// TIA Portal V20 export
VAR_GLOBAL   // PLC tag table "COGNEX_ETIKETA"
   "COG_ETIKETA_COG_ETIKETA_is3800-TriggerEnable" AT %Q2.0 : Bool;
   "COG_ETIKETA_COG_ETIKETA_is3800-Trigger" AT %Q2.1 : Bool;
   "COG_ETIKETA_is3800-ClearExposureComplete" AT %Q2.2 : Bool;
   "COG_ETIKETA_is3800-Set Offline" AT %Q2.7 : Bool;
   "COG_ETIKETA_is3800-TriggerReady" AT %I2.0 : Bool;
   "COG_ETIKETA_is3800-TriggerAck" AT %I2.1 : Bool;
   "COG_ETIKETA_is3800-ExposureComplete" AT %I2.2 : Bool;
   "COG_ETIKETA_is3800-AcquCOG_ETIKETA_isitionError" AT %I2.3 : Bool;
   "COG_ETIKETA_is3800-Offline Reason" AT %I2.4 : Bool;
   "COG_ETIKETA_is3800-Offline Reason(1)" AT %I2.5 : Bool;
   "COG_ETIKETA_is3800-Offline Reason(2)" AT %I2.6 : Bool;
   "COG_ETIKETA_is3800-Online" AT %I2.7 : Bool;
   "COG_ETIKETA_is3800-AcquCOG_ETIKETA_isitionID" AT %IW4 : Int;
   "COG_ETIKETA_is3800-BufferResultsEnable" AT %Q3.0 : Bool;
   "COG_ETIKETA_is3800-InspectionResultsAck" AT %Q3.1 : Bool;
   "COG_ETIKETA_is3800-SetUserData" AT %Q3.2 : Bool;
   "COG_ETIKETA_is3800-ExecuteCommand/JobLoad" AT %Q3.3 : Bool;
   "COG_ETIKETA_is3800-ClearError" AT %Q3.7 : Bool;
   "COG_ETIKETA_is3800-Reserved" AT %I10.0 : Bool;
   "COG_ETIKETA_is3800-InspectionCompleted" AT %I10.1 : Bool;
   "COG_ETIKETA_is3800-ResultsBufferOverrun" AT %I10.2 : Bool;
   "COG_ETIKETA_is3800-ResultsValid" AT %I10.3 : Bool;
   "COG_ETIKETA_is3800-CommandExecuting" AT %I10.4 : Bool;
   "COG_ETIKETA_is3800-CommandCompleted" AT %I10.5 : Bool;
   "COG_ETIKETA_is3800-CommandFailed" AT %I10.6 : Bool;
   "COG_ETIKETA_is3800-SetUserDataAck" AT %I10.7 : Bool;
   "COG_ETIKETA_is3800-ResultsPassed (Job)" AT %I11.0 : Bool;
   "COG_ETIKETA_is3800-SystemValidated" AT %I11.1 : Bool;
   "COG_ETIKETA_is3800-Error" AT %I11.7 : Bool;
   "COG_ETIKETA_is3800-ErrorCode" AT %IW12 : Word;
   "COG_ETIKETA_is3800-CommandID" AT %QW64 : Word;
   "COG_ETIKETA_is3800-Current Job ID" AT %IW68 : Word;
   "COG_ETIKETA_is3800-CommandResultCode" AT %IW70 : Word;
   "COG_ETIKETA_is3800-ExternalEvent[0]" AT %Q4.0 : Bool;
   "COG_ETIKETA_is3800-ExternalEvent[1]" AT %Q4.1 : Bool;
   "COG_ETIKETA_is3800-ExternalEvent[2]" AT %Q4.2 : Bool;
   "COG_ETIKETA_is3800-ExternalEvent[3]" AT %Q4.3 : Bool;
   "COG_ETIKETA_is3800-ExternalEvent[4]" AT %Q4.4 : Bool;
   "COG_ETIKETA_is3800-ExternalEvent[5]" AT %Q4.5 : Bool;
   "COG_ETIKETA_is3800-ExternalEvent[6]" AT %Q4.6 : Bool;
   "COG_ETIKETA_is3800-ExternalEvent[7]" AT %Q4.7 : Bool;
   "COG_ETIKETA_is3800-ExternalEventAck[0]" AT %I6.0 : Bool;
   "COG_ETIKETA_is3800-ExternalEventAck[1]" AT %I6.1 : Bool;
   "COG_ETIKETA_is3800-ExternalEventAck[2]" AT %I6.2 : Bool;
   "COG_ETIKETA_is3800-ExternalEventAck[3]" AT %I6.3 : Bool;
   "COG_ETIKETA_is3800-ExternalEventAck[4]" AT %I6.4 : Bool;
   "COG_ETIKETA_is3800-ExternalEventAck[5]" AT %I6.5 : Bool;
   "COG_ETIKETA_is3800-ExternalEventAck[6]" AT %I6.6 : Bool;
   "COG_ETIKETA_is3800-ExternalEventAck[7]" AT %I6.7 : Bool;
   "COG_ETIKETA_is3800-UserData[0]" AT %QB66 : Byte;
   "COG_ETIKETA_is3800-UserData[1]" AT %QB67 : Byte;
   "COG_ETIKETA_is3800-UserData[2]" AT %QB68 : Byte;
   "COG_ETIKETA_is3800-UserData[3]" AT %QB69 : Byte;
   "COG_ETIKETA_is3800-UserData[4]" AT %QB70 : Byte;
   "COG_ETIKETA_is3800-UserData[5]" AT %QB71 : Byte;
   "COG_ETIKETA_is3800-UserData[6]" AT %QB72 : Byte;
   "COG_ETIKETA_is3800-UserData[7]" AT %QB73 : Byte;
   "COG_ETIKETA_is3800-UserData[8]" AT %QB74 : Byte;
   "COG_ETIKETA_is3800-UserData[9]" AT %QB75 : Byte;
   "COG_ETIKETA_is3800-UserData[10]" AT %QB76 : Byte;
   "COG_ETIKETA_is3800-UserData[11]" AT %QB77 : Byte;
   "COG_ETIKETA_is3800-UserData[12]" AT %QB78 : Byte;
   "COG_ETIKETA_is3800-UserData[13]" AT %QB79 : Byte;
   "COG_ETIKETA_is3800-UserData[14]" AT %QB80 : Byte;
   "COG_ETIKETA_is3800-UserData[15]" AT %QB81 : Byte;
   "COG_ETIKETA_is3800-InspectionID" AT %IW72 : Word;
   "COG_ETIKETA_is3800-InspectionResultsCode" AT %IW74 : Int;
   "COG_ETIKETA_is3800-InspectionResults_0" AT %IB76 : Byte;
   "COG_ETIKETA_is3800-InspectionResults_1" AT %IB77 : Byte;
   "COG_ETIKETA_is3800-InspectionResults_2" AT %IB78 : Byte;
   "COG_ETIKETA_is3800-InspectionResults_3" AT %IB79 : Byte;
   "COG_ETIKETA_is3800-InspectionResults_4" AT %IB80 : Byte;
   "COG_ETIKETA_is3800-InspectionResults_5" AT %IB81 : Byte;
   "COG_ETIKETA_is3800-InspectionResults_6" AT %IB82 : Byte;
   "COG_ETIKETA_is3800-InspectionResults_7" AT %IB83 : Byte;
   "COG_ETIKETA_is3800-InspectionResults_8" AT %IB84 : Byte;
   "COG_ETIKETA_is3800-InspectionResults_9" AT %IB85 : Byte;
   "COG_ETIKETA_is3800-InspectionResults_10" AT %IB86 : Byte;
   "COG_ETIKETA_is3800-InspectionResults_11" AT %IB87 : Byte;
   "COG_ETIKETA_is3800-InspectionResults_12" AT %IB88 : Byte;
   "COG_ETIKETA_is3800-InspectionResults_13" AT %IB89 : Byte;
   "COG_ETIKETA_is3800-InspectionResults_14" AT %IB90 : Byte;
   "COG_ETIKETA_is3800-InspectionResults_15" AT %IB91 : Byte;
   "COG_ETIKETA_is3800-InspectionResults_16" AT %IB92 : Byte;
   "COG_ETIKETA_is3800-InspectionResults_17" AT %IB93 : Byte;
   "COG_ETIKETA_is3800-InspectionResults_18" AT %IB94 : Byte;
   "COG_ETIKETA_is3800-InspectionResults_19" AT %IB95 : Byte;
   "COG_ETIKETA_is3800-InspectionResults_20" AT %IB96 : Byte;
   "COG_ETIKETA_is3800-InspectionResults_21" AT %IB97 : Byte;
   "COG_ETIKETA_is3800-InspectionResults_22" AT %IB98 : Byte;
   "COG_ETIKETA_is3800-InspectionResults_23" AT %IB99 : Byte;
   "COG_ETIKETA_is3800-InspectionResults_24" AT %IB100 : Byte;
   "COG_ETIKETA_is3800-InspectionResults_25" AT %IB101 : Byte;
   "COG_ETIKETA_is3800-InspectionResults_26" AT %IB102 : Byte;
   "COG_ETIKETA_is3800-InspectionResults_27" AT %IB103 : Byte;
   "COG_ETIKETA_is3800-InspectionResults_28" AT %IB104 : Byte;
   "COG_ETIKETA_is3800-InspectionResults_29" AT %IB105 : Byte;
   "COG_ETIKETA_is3800-InspectionResults_30" AT %IB106 : Byte;
   "COG_ETIKETA_is3800-InspectionResults_31" AT %IB107 : Byte;
   "COG_ETIKETA_is3800-InspectionResults_32" AT %IB108 : Byte;
   "COG_ETIKETA_is3800-InspectionResults_33" AT %IB109 : Byte;
   "COG_ETIKETA_is3800-InspectionResults_34" AT %IB110 : Byte;
   "COG_ETIKETA_is3800-InspectionResults_35" AT %IB111 : Byte;
   "COG_ETIKETA_is3800-InspectionResults_36" AT %IB112 : Byte;
   "COG_ETIKETA_is3800-InspectionResults_37" AT %IB113 : Byte;
   "COG_ETIKETA_is3800-InspectionResults_38" AT %IB114 : Byte;
   "COG_ETIKETA_is3800-InspectionResults_39" AT %IB115 : Byte;
   "COG_ETIKETA_is3800-InspectionResults_40" AT %IB116 : Byte;
   "COG_ETIKETA_is3800-InspectionResults_41" AT %IB117 : Byte;
   "COG_ETIKETA_is3800-InspectionResults_42" AT %IB118 : Byte;
   "COG_ETIKETA_is3800-InspectionResults_43" AT %IB119 : Byte;
   "COG_ETIKETA_is3800-InspectionResults_44" AT %IB120 : Byte;
   "COG_ETIKETA_is3800-InspectionResults_45" AT %IB121 : Byte;
   "COG_ETIKETA_is3800-InspectionResults_46" AT %IB122 : Byte;
   "COG_ETIKETA_is3800-InspectionResults_47" AT %IB123 : Byte;
   "COG_ETIKETA_is3800-InspectionResults_48" AT %IB124 : Byte;
   "COG_ETIKETA_is3800-InspectionResults_49" AT %IB125 : Byte;
   "COG_ETIKETA_is3800-InspectionResults_50" AT %IB126 : Byte;
   "COG_ETIKETA_is3800-InspectionResults_51" AT %IB127 : Byte;
   "COG_ETIKETA_is3800-InspectionResults_52" AT %IB128 : Byte;
   "COG_ETIKETA_is3800-InspectionResults_53" AT %IB129 : Byte;
   "COG_ETIKETA_is3800-InspectionResults_54" AT %IB130 : Byte;
   "COG_ETIKETA_is3800-InspectionResults_55" AT %IB131 : Byte;
   "COG_ETIKETA_is3800-InspectionResults_56" AT %IB132 : Byte;
   "COG_ETIKETA_is3800-InspectionResults_57" AT %IB133 : Byte;
   "COG_ETIKETA_is3800-InspectionResults_58" AT %IB134 : Byte;
   "COG_ETIKETA_is3800-InspectionResults_59" AT %IB135 : Byte;
   "COG_ETIKETA_is3800-InspectionResults_60" AT %IB136 : Byte;
   "COG_ETIKETA_is3800-InspectionResults_61" AT %IB137 : Byte;
   "COG_ETIKETA_is3800-InspectionResults_62" AT %IB138 : Byte;
   "COG_ETIKETA_is3800-InspectionResults_63" AT %IB139 : Byte;
   "COG_ETIKETA_is3800-InspectionResults_64" AT %IB140 : Byte;
   "COG_ETIKETA_is3800-InspectionResults_65" AT %IB141 : Byte;
   "COG_ETIKETA_is3800-InspectionResults_66" AT %IB142 : Byte;
   "COG_ETIKETA_is3800-InspectionResults_67" AT %IB143 : Byte;
   "COG_ETIKETA_is3800-InspectionResults_68" AT %IB144 : Byte;
   "COG_ETIKETA_is3800-InspectionResults_69" AT %IB145 : Byte;
   "COG_ETIKETA_is3800-InspectionResults_70" AT %IB146 : Byte;
   "COG_ETIKETA_is3800-InspectionResults_71" AT %IB147 : Byte;
   "COG_ETIKETA_is3800-InspectionResults_72" AT %IB148 : Byte;
   "COG_ETIKETA_is3800-InspectionResults_73" AT %IB149 : Byte;
   "COG_ETIKETA_is3800-InspectionResults_74" AT %IB150 : Byte;
   "COG_ETIKETA_is3800-InspectionResults_75" AT %IB151 : Byte;
   "COG_ETIKETA_is3800-InspectionResults_76" AT %IB152 : Byte;
   "COG_ETIKETA_is3800-InspectionResults_77" AT %IB153 : Byte;
   "COG_ETIKETA_is3800-InspectionResults_78" AT %IB154 : Byte;
   "COG_ETIKETA_is3800-InspectionResults_79" AT %IB155 : Byte;
   "COG_ETIKETA_is3800-InspectionResults_80" AT %IB156 : Byte;
   "COG_ETIKETA_is3800-InspectionResults_81" AT %IB157 : Byte;
   "COG_ETIKETA_is3800-InspectionResults_82" AT %IB158 : Byte;
   "COG_ETIKETA_is3800-InspectionResults_83" AT %IB159 : Byte;
   "COG_ETIKETA_is3800-InspectionResults_84" AT %IB160 : Byte;
   "COG_ETIKETA_is3800-InspectionResults_85" AT %IB164 : Byte;
   "COG_ETIKETA_is3800-InspectionResults_86" AT %IB165 : Byte;
   "COG_ETIKETA_is3800-InspectionResults_87" AT %IB166 : Byte;
   "COG_ETIKETA_is3800-InspectionResults_88" AT %IB167 : Byte;
   "COG_ETIKETA_is3800-InspectionResults_89" AT %IB168 : Byte;
   "COG_ETIKETA_is3800-InspectionResults_90" AT %IB169 : Byte;
   "COG_ETIKETA_is3800-InspectionResults_91" AT %IB170 : Byte;
   "COG_ETIKETA_is3800-InspectionResults_92" AT %IB171 : Byte;
   "COG_ETIKETA_is3800-InspectionResults_93" AT %IB172 : Byte;
   "COG_ETIKETA_is3800-InspectionResults_94" AT %IB173 : Byte;
   "COG_ETIKETA_is3800-InspectionResults_95" AT %IB174 : Byte;
   "COG_ETIKETA_is3800-InspectionResults_96" AT %IB175 : Byte;
   "COG_ETIKETA_is3800-InspectionResults_97" AT %IB176 : Byte;
   "COG_ETIKETA_is3800-InspectionResults_98" AT %IB177 : Byte;
   "COG_ETIKETA_is3800-InspectionResults_99" AT %IB178 : Byte;
   "COG_ETIKETA_is3800-InspectionResults_100" AT %IB179 : Byte;
END_VAR
